(* IEC 61131-3 sources: PLC_ST_Auto/examples, 21 files *)

(* ---- aoi_l5x.st ---- *)
(* M35:自訂 FUNCTION_BLOCK → Rockwell L5X Add-On Instruction 匯出範例 *)
FUNCTION_BLOCK Latch
VAR_INPUT set : BOOL; rst : BOOL; END_VAR
VAR_OUTPUT q : BOOL; n : INT; END_VAR
VAR rt : R_TRIG; END_VAR
rt(CLK := set);
IF rt.Q THEN n := n + 1; END_IF;
IF set THEN q := TRUE; END_IF;
IF rst THEN q := FALSE; END_IF;
END_FUNCTION_BLOCK

FUNCTION_BLOCK Accum
VAR_INPUT add : DINT := 1; go : BOOL; END_VAR
VAR_IN_OUT shared : DINT; END_VAR
VAR_OUTPUT total : DINT; END_VAR
VAR CONSTANT LAST : INT := 3; END_VAR
VAR i : INT; inner : Latch; buf : ARRAY[0..3] OF DINT := [1, 2, 3, 4]; END_VAR
inner(set := go, rst := FALSE);
IF inner.q THEN
  total := 0;
  FOR i := 0 TO LAST DO
    buf[i] := buf[i] + add;
    total := total + buf[i];
  END_FOR;
  shared := shared + total;
END_IF;
END_FUNCTION_BLOCK

PROGRAM Main
VAR_INPUT start : BOOL; stop : BOOL; END_VAR
VAR_OUTPUT pump : BOOL; starts : INT; sum : DINT; END_VAR
VAR l1 : Latch; acc : Accum; pool : DINT; END_VAR
l1(set := start, rst := stop, q => pump);
starts := l1.n;
IF start THEN
  acc(add := 10, go := start, shared := pool, total => sum);
END_IF;
END_PROGRAM

(* ---- array_inout.st ---- *)
(* M36:整個陣列傳入 VAR_IN_OUT / VAR_INPUT、陣列整體賦值 *)
FUNCTION SumAndDouble : DINT
VAR_IN_OUT data : ARRAY[1..5] OF INT; END_VAR
VAR i : INT; END_VAR
SumAndDouble := 0;
FOR i := 1 TO 5 DO
  SumAndDouble := SumAndDouble + data[i];
  data[i] := data[i] * 2;
END_FOR;
END_FUNCTION

FUNCTION_BLOCK ShiftReg
VAR_INPUT nv : INT; END_VAR
VAR_IN_OUT buf : ARRAY[0..4] OF INT; END_VAR
VAR k : INT; END_VAR
FOR k := 4 TO 1 BY -1 DO
  buf[k] := buf[k - 1];
END_FOR;
buf[0] := nv;
END_FUNCTION_BLOCK

FUNCTION MaxOf : INT
VAR_INPUT v : ARRAY[0..4] OF INT; END_VAR
VAR i : INT; END_VAR
MaxOf := v[0];
FOR i := 1 TO 4 DO
  IF v[i] > MaxOf THEN MaxOf := v[i]; END_IF;
END_FOR;
END_FUNCTION

PROGRAM Main
VAR_INPUT
  sample : INT;
END_VAR
VAR
  hist : ARRAY[0..4] OF INT;
  snap : ARRAY[0..4] OF INT;
  sh : ShiftReg;
  peak : INT;
END_VAR
sh(nv := sample, buf := hist);
snap := hist;
peak := MaxOf(snap);
END_PROGRAM

(* ---- global_vars.st ---- *)
(* M43 範例:VAR_GLOBAL / VAR_EXTERNAL(CODESYS GVL 寫法)
   兩條輸送帶共用全域計數 g_count、全域上限 G_LIMIT(常數)與全域停止旗標 g_stop *)
VAR_GLOBAL CONSTANT
    G_LIMIT : INT := 5;
END_VAR
VAR_GLOBAL
    g_count : INT := 0;
    g_stop : BOOL;
    g_log : ARRAY[0..3] OF INT;
END_VAR

FUNCTION_BLOCK FB_Counter
VAR_INPUT
    pulse : BOOL;
END_VAR
VAR_EXTERNAL
    g_count : INT;
    g_stop : BOOL;
    g_log : ARRAY[0..3] OF INT;
END_VAR
VAR_EXTERNAL CONSTANT
    G_LIMIT : INT;
END_VAR
VAR
    edge : R_TRIG;
    mine : INT;
END_VAR
edge(CLK := pulse);
IF edge.Q AND NOT g_stop THEN
    g_count := g_count + 1;
    mine := mine + 1;
    g_log[g_count MOD 4] := mine;
END_IF;
g_stop := g_count >= G_LIMIT;
END_FUNCTION_BLOCK

FUNCTION Remaining : INT
VAR_EXTERNAL
    g_count : INT;
END_VAR
VAR_EXTERNAL CONSTANT
    G_LIMIT : INT;
END_VAR
Remaining := G_LIMIT - g_count;
END_FUNCTION

PROGRAM Main
VAR_INPUT
    sensorA : BOOL;
    sensorB : BOOL;
    reset : BOOL;
END_VAR
VAR_OUTPUT
    full : BOOL;
    remain : INT;
END_VAR
VAR
    cA : FB_Counter;
    cB : FB_Counter;
END_VAR
cA(pulse := sensorA);
cB(pulse := sensorB);
IF reset THEN
    g_count := 0;
END_IF;
full := g_stop;
remain := Remaining();
END_PROGRAM

(* ---- inout.st ---- *)
FUNCTION Bump : INT
VAR_INPUT step : INT; END_VAR
VAR_IN_OUT v : INT; END_VAR
v := v + step;
Bump := v;
END_FUNCTION

FUNCTION_BLOCK Acc
VAR_INPUT d : INT; END_VAR
VAR_IN_OUT total : INT; END_VAR
total := total + d;
END_FUNCTION_BLOCK

PROGRAM P
VAR
  x : INT := 1; r : INT; y : INT := 10;
  a1 : Acc;
END_VAR
r := Bump(step := 2, v := x);
a1(d := 5, total := y);
END_PROGRAM

(* ---- recipe_slots.st ---- *)
(* 配方槽:ARRAY OF STRUCT,且 STRUCT 內含 ARRAY 欄位(M41) *)
TYPE Recipe : STRUCT
  setp : ARRAY[1..3] OF INT := [100, 200, 300];
  hold : ARRAY[1..3] OF TIME;
  name : STRING := 'empty';
END_STRUCT
END_TYPE

FUNCTION_BLOCK StepRunner
VAR_INPUT run : BOOL; END_VAR
VAR_IN_OUT sp : ARRAY[1..3] OF INT; END_VAR
VAR_OUTPUT total : INT; END_VAR
VAR i : INT; END_VAR
total := 0;
FOR i := 1 TO 3 DO
  IF run THEN sp[i] := sp[i] + 1; END_IF;
  total := total + sp[i];
END_FOR;
END_FUNCTION_BLOCK

PROGRAM Main
VAR_INPUT
  slot : INT := 1;
  bump : BOOL;
  save : BOOL;
END_VAR
VAR_OUTPUT
  active : ARRAY[1..3] OF INT;
  sum : INT;
END_VAR
VAR
  slots : ARRAY[1..3] OF Recipe := [(name := 'A'), (setp := [10, 20, 30], name := 'B')];
  work : Recipe;
  runner : StepRunner;
  k : INT;
  n : INT;
END_VAR
n := LIMIT(1, slot, 3);
work := slots[n];                       (* 整個元素複製到單一 STRUCT *)
active := slots[n].setp;                (* 元素的陣列欄位整體讀出 *)
runner(run := bump, sp := slots[n].setp, total => sum);   (* VAR_IN_OUT 寫回元素的陣列欄位 *)
IF save THEN
  FOR k := 1 TO 3 DO
    slots[3].setp[k] := slots[n].setp[k] * 2;
  END_FOR;
  slots[3].name := 'copy';
END_IF;
END_PROGRAM

(* ---- userpou_export.st ---- *)
(* M33:自訂 FUNCTION / FUNCTION_BLOCK 匯出範例(PLCopen XML、Siemens SCL) *)
FUNCTION Scale : REAL
VAR_INPUT raw : INT; hi : REAL; END_VAR
VAR k : REAL := 100.0; END_VAR
Scale := INT_TO_REAL(raw) * hi / k;
END_FUNCTION

FUNCTION Clamp : INT
VAR_INPUT x : INT; lo : INT; top : INT; END_VAR
IF x > top THEN
  Clamp := top;
  RETURN;
END_IF;
Clamp := MAX(x, lo);
END_FUNCTION

FUNCTION_BLOCK Latch
VAR_INPUT set : BOOL; rst : BOOL; END_VAR
VAR_OUTPUT q : BOOL; n : INT; END_VAR
VAR rt : R_TRIG; END_VAR
rt(CLK := set);
IF rt.Q THEN n := n + 1; END_IF;
IF set THEN q := TRUE; END_IF;
IF rst THEN q := FALSE; END_IF;
END_FUNCTION_BLOCK

PROGRAM Main
VAR_INPUT start : BOOL; stop : BOOL; level_raw : INT; END_VAR
VAR_OUTPUT pump : BOOL; level : REAL; starts : INT; duty : INT; END_VAR
VAR l1 : Latch; msg : STRING := 'Clamp(1, 2)'; END_VAR
level := Scale(level_raw, 200.0);            (* 位置引數 *)
duty := Clamp(REAL_TO_INT(Scale(raw := level_raw, hi := 100.0)), 0, 80);
l1(set := start, rst := stop);
pump := l1.q;
starts := l1.n;
END_PROGRAM

(* ---- literals_m31.st ---- *)
PROGRAM literals
VAR
    a : INT; b : REAL; t : TIME; c : INT; h : DINT; f : BOOL;
    m : ARRAY[0..4] OF INT := [2(1), 3(0)];
END_VAR
a := INT#5 + 16#FF + 2#1010 + 1_000;
b := INT_TO_REAL(a) + REAL#1.5;
t := INT_TO_TIME(250);
c := TIME_TO_INT(t) + REAL_TO_INT(2.6);
h := 8#17;
f := BOOL#1;
END_PROGRAM

(* ---- m32_escape_round.st ---- *)
PROGRAM m32
VAR
  msg : STRING := 'it$'s $$5$N';
  n : INT;
  r : REAL := 2.5;
  rounded : INT;
  cnt : INT;
END_VAR
n := LEN(msg);
rounded := r;            (* 2.5 -> 3 (遠離零) *)
FOR cnt := 0 TO 10 DO
  IF cnt = 4 THEN EXIT; END_IF
END_FOR
END_PROGRAM

(* ---- matrix.st ---- *)
PROGRAM Matrix
VAR
  m : ARRAY[1..2, 1..3] OF INT := [1, 2, 3, 4, 5, 6];
  i : INT := 1;
  j : INT := 1;
  total : INT;
END_VAR
total := 0;
FOR i := 1 TO 2 DO
  FOR j := 1 TO 3 DO
    total := total + m[i, j];
  END_FOR;
END_FOR;
m[2, 3] := m[2, 3] + 1;
END_PROGRAM

(* ---- motor.st ---- *)
PROGRAM Motor
VAR_INPUT start : BOOL; stop : BOOL; END_VAR
VAR_OUTPUT motor : BOOL; END_VAR
VAR t : TON; cnt : INT; END_VAR
IF start AND NOT stop THEN motor := TRUE; END_IF;
IF stop THEN motor := FALSE; END_IF;
t(IN := motor, PT := T#500ms);
IF t.Q THEN cnt := cnt + 1; END_IF;
END_PROGRAM

(* ---- qualifiers_m34.st ---- *)
(* M34:VAR CONSTANT / RETAIN / VAR_TEMP 與直接位址 AT %I/%Q/%M *)
PROGRAM Conveyor
VAR CONSTANT
  N : INT := 4;              (* 站數 *)
  MAX_COUNT : DINT := 1000;
END_VAR
VAR RETAIN
  total : DINT;              (* 斷電保持的累計數量 *)
END_VAR
VAR_TEMP
  i : INT;
  sum : INT := 0;
END_VAR
VAR
  start AT %IX0.0 : BOOL;
  sensor AT %IX0.1 : BOOL;
  motor AT %QX0.0 : BOOL;
  speed AT %QW2 : INT;
  full AT %MX1.0 : BOOL;
  slots : ARRAY[0..N - 1] OF INT := [1, 2, 3, 4];
  edge : R_TRIG;
  batch : DINT;
END_VAR
edge(CLK := sensor);
IF edge.Q AND total < MAX_COUNT THEN
  total := total + 1;
  batch := batch + 1;
END_IF;
FOR i := 0 TO N - 1 DO
  sum := sum + slots[i];
END_FOR;
motor := start AND NOT full;
full := total >= MAX_COUNT;
speed := sum * 10;   // 'start' in a string or (* start *) comment stays untouched
END_PROGRAM

(* ---- review_m29.st ---- *)
(* M29 審查修正示範:8 個 BOOL、字串含 // ; (*、陣列邊界運算式、實例陣列初值 *)
TYPE Flags : STRUCT
  f0, f1, f2, f3, f4, f5, f6, f7 : BOOL;
  url : STRING := 'http://host/a;b';
  buf : ARRAY[0..2+1] OF INT := [1, 2];
END_STRUCT END_TYPE
PROGRAM Demo
VAR
  a : Flags := (buf := [10, 20, 30, 40]);
  b : Flags;
  hist : ARRAY[0..(1+1)*2] OF INT;
  i : INT;
  sum : INT;
END_VAR
a.f7 := TRUE;
sum := 0;
FOR i := 0 TO 3 DO sum := sum + a.buf[i] + b.buf[i]; END_FOR
hist[4] := sum;
END_PROGRAM

(* ---- shared_memory.st ---- *)
(* M37:直接位址共用記憶體。
   %IB0 是整個輸入位元組,start / stop 是其中的位元;%MW0 狀態字與 %MX 旗標共用位元組。
   位元組順序依 profile:IEC/CODESYS 為 little-endian(%MX0.0 = %MW0 bit 0),
   Siemens 為 big-endian(%M0.0 = %MW0 bit 8,%M1.0 = bit 0)。 *)
PROGRAM SharedMem
VAR
    inByte  AT %IB0   : BYTE;     (* 整個輸入位元組:可一次強制 8 個輸入 *)
    start   AT %IX0.0 : BOOL;
    stop    AT %IX0.1 : BOOL;
    status  AT %MW0   : WORD;     (* 狀態字,例如送到 HMI *)
    running AT %MX0.0 : BOOL;     (* IEC:status 的 bit 0;Siemens:bit 8 *)
    alarm   AT %MX1.7 : BOOL;     (* IEC:status 的 bit 15;Siemens:bit 7 *)
    motor   AT %QX0.0 : BOOL;
    outByte AT %QB0   : BYTE;
END_VAR
IF start AND NOT stop THEN
    running := TRUE;
ELSIF stop THEN
    running := FALSE;
END_IF;
alarm := start AND stop;
motor := running;
END_PROGRAM

(* ---- struct.st ---- *)
TYPE Motor : STRUCT
  speed : INT := 10;
  run : BOOL;
END_STRUCT END_TYPE
TYPE Line : STRUCT
  m : Motor;
  count : DINT;
END_STRUCT END_TYPE
PROGRAM P
VAR
  a : Motor := (speed := 50);
  l : Line := (count := 3, m := (speed := 7));
  t : TON;
END_VAR
a.run := a.speed > 20;
l.m.speed := l.m.speed + 1;
l.count := l.count + a.speed;
END_PROGRAM

(* ---- struct_array.st ---- *)
TYPE Motor : STRUCT
  speed : INT := 10;
  run : BOOL;
END_STRUCT END_TYPE
PROGRAM P
VAR
  ms : ARRAY[1..3] OF Motor;
  i : INT;
  total : INT;
END_VAR
total := 0;
FOR i := 1 TO 3 DO
  ms[i].speed := ms[i].speed + i;
  ms[i].run := ms[i].speed > 11;
  total := total + ms[i].speed;
END_FOR;
END_PROGRAM

(* ---- struct_arrfield.st ---- *)
TYPE Recipe : STRUCT
  id : INT := 5;
  steps : ARRAY[0..3] OF INT := [10, 20];
  grid : ARRAY[1..2, 1..2] OF REAL;
END_STRUCT END_TYPE
PROGRAM P
VAR
  r, backup : Recipe;
  i : INT;
  total : INT;
END_VAR
FOR i := 0 TO 3 DO r.steps[i] := r.steps[i] + i; END_FOR
r.grid[2, 1] := 2.5;
backup := r;
r.steps[0] := 99;
total := backup.steps[0] + backup.steps[3] + r.id;
END_PROGRAM

(* ---- struct_copy.st ---- *)
TYPE Motor : STRUCT
  speed : INT := 10;
  run : BOOL;
END_STRUCT END_TYPE
TYPE Line : STRUCT
  m : Motor;
  count : DINT;
END_STRUCT END_TYPE
PROGRAM P
VAR
  a : Motor := (speed := 50);
  b : Motor;
  l : Line;
END_VAR
a.run := TRUE;
b := a;          (* whole-STRUCT copy *)
l.m := b;        (* nested STRUCT copy *)
l.count := l.count + 1;
a.speed := a.speed + 1;
END_PROGRAM

(* ---- struct_elem.st ---- *)
TYPE Motor : STRUCT
  speed : INT := 10;
  run : BOOL;
END_STRUCT END_TYPE
PROGRAM P
VAR
  ms : ARRAY[1..3] OF Motor := [(speed := 100, run := TRUE), (speed := 200)];
  tmp : Motor;
  best : INT;
END_VAR
tmp := ms[1];
ms[3] := ms[2];
ms[2] := tmp;
best := ms[3].speed;
END_PROGRAM

(* ---- struct_export.st ---- *)
TYPE Motor : STRUCT
  speed : INT := 10;
  run : BOOL;
END_STRUCT END_TYPE
PROGRAM P
VAR
  ms : ARRAY[1..3] OF Motor := [(speed := 100, run := TRUE), (speed := 200)];
  tmp : Motor;
  best : INT;
END_VAR
tmp := ms[1];
ms[3] := ms[2];
ms[2] := tmp;
best := ms[3].speed;
END_PROGRAM

(* ---- struct_gx_sysmac.st ---- *)
(* M42:TYPE STRUCT 匯出 GX Works3 / Sysmac Studio 範例(巢狀 STRUCT、陣列欄位、ARRAY OF STRUCT 初值) *)
TYPE Pt : STRUCT
  x : INT := 1;
  y : INT;
END_STRUCT END_TYPE
TYPE Axis : STRUCT
  home : Pt;
  pos : ARRAY[0..1] OF INT := [0, 0];
  name : STRING := 'axis';
  ready : BOOL;
END_STRUCT END_TYPE
PROGRAM P
VAR_INPUT
  start : BOOL;
END_VAR
VAR_OUTPUT
  sum : INT;
END_VAR
VAR
  ax : Axis := (home := (x := 5, y := 6), name := 'X, main');
  marks : ARRAY[1..3] OF Pt := [(x := 10), 2((y := 20))];
END_VAR
IF start THEN
  ax.pos[1] := ax.pos[1] + 1;
  ax.ready := ax.pos[1] >= 3;
END_IF;
sum := ax.home.x + ax.home.y + marks[1].x + marks[3].y + ax.pos[1];
END_PROGRAM

(* ---- struct_l5x.st ---- *)
TYPE Motor : STRUCT
  speed : INT;
  run : BOOL;
END_STRUCT END_TYPE
PROGRAM P
VAR
  ms : ARRAY[0..2] OF Motor;
  best : INT;
END_VAR
ms[1].speed := 200;
ms[1].run := TRUE;
best := ms[1].speed;
END_PROGRAM
